Universal Robots PolyScope program: Renee_AI.urp

Program Renee_AI (installation=default directory=/ursim/programs createdIn=5.26.0 lastSavedIn=5.26.1 robotSerialNumber=20195599999)
Calibrated DH parameters: a=[0, -0.425, -0.3922, 0, 0, 0]; d=[0.1625, 0, 0, 0.1333, 0.0997, 0.0996]; alpha=[1.570796, 0, 0, 1.570796, -1.570796, 0]; deltaTheta=[0, 0, 0, 0, 0, 0]
InitVariablesNode
Robot Program (runOnlyOnce=true)
  var_1 := get_actual_tcp_pose()
  MoveJ speed 60 deg/s, acceleration 80 deg/s^2 (useActiveTCP=true optimoveEnabled=false optiMoveSpeed=0.3 optiMoveAcceleration=0.09) feature=Base
    Waypoint Variable (Variable): variable=var_1
  MoveJ speed 60 deg/s, acceleration 80 deg/s^2 (useActiveTCP=true positionType=JointAngles optimoveEnabled=false optiMoveSpeed=0.3 optiMoveAcceleration=0.09) feature=Base
    Waypoint Waypoint_1: TCP in base x=202.351 y=489.879 z=593.238 mm, rx=-1.5225 ry=0.5256 rz=-0.412 rad; joints [-127.677, -86.227, 99.579, -191.944, -86.567, 3.764] deg
  Script file /ursim/programs/generated_task.script
    | def inspection_program():
    |   # T_base_cam as a UR pose (position + axis-angle rotation vector)
    |   # Derived from the 4x4 transformation matrix T_base_cam
    |   global T_base_cam = p[0.352728458264352, -0.21258760881184183, 0.11788934094986696, -1.538543, 0.024168, 0.017202]
    | 
    |   # Offset to apply in camera frame: -0.4 m in camera X
    |   global x_offset = -0.40
    | 
    |   # Movement parameters (conservative for inspection)
    |   global accel = 0.3
    |   global vel = 0.05
    | 
    |   # Compute the first waypoint pose
    |   local first_wp = pose_trans(T_base_cam, p[0.335 + x_offset, 0.143, 0.57, 0, 0, 0])
    | 
    |   # Use movej to safely approach the first waypoint (avoids protective stop)
    |   movej(first_wp, a=1.0, v=0.5)
    |   sleep(1.0)
    | 
    |   # --- Waypoint 2: top_tube_front ---
    |   movel(pose_trans(T_base_cam, p[0.381 + x_offset, 0.116, 0.57, 0, 0, 0]), a=accel, v=vel)
    |   sleep(1.0)
    | 
    |   # --- Waypoint 3: top_tube_rear ---
    |   movel(pose_trans(T_base_cam, p[0.65 + x_offset, 0.131, 0.57, 0, 0, 0]), a=accel, v=vel)
    |   sleep(1.0)
    | 
    |   # --- Waypoint 4: seat_post_clamp ---
    |   movel(pose_trans(T_base_cam, p[0.68 + x_offset, 0.11, 0.57, 0, 0, 0]), a=accel, v=vel)
    |   sleep(1.0)
    | 
    |   # --- Waypoint 5: seat_tube_lower ---
    |   movel(pose_trans(T_base_cam, p[0.627 + x_offset, 0.462, 0.57, 0, 0, 0]), a=accel, v=vel)
    |   sleep(1.0)
    | 
    |   # --- Waypoint 6: bottom_bracket ---
    |   movel(pose_trans(T_base_cam, p[0.615 + x_offset, 0.609, 0.57, 0, 0, 0]), a=accel, v=vel)
    |   sleep(1.0)
    | 
    |   # --- Waypoint 7: chainstay_front ---
    |   movel(pose_trans(T_base_cam, p[0.701 + x_offset, 0.609, 0.57, 0, 0, 0]), a=accel, v=vel)
    |   sleep(1.0)
    | 
    |   # --- Waypoint 8: rear_dropout ---
    |   movel(pose_trans(T_base_cam, p[0.888 + x_offset, 0.586, 0.57, 0, 0, 0]), a=accel, v=vel)
    |   sleep(1.0)
    | 
    |   # --- Waypoint 9: seatstay_upper ---
    |   movel(pose_trans(T_base_cam, p[0.736 + x_offset, 0.308, 0.57, 0, 0, 0]), a=accel, v=vel)
    |   sleep(1.0)
    | 
    |   # --- Waypoint 10: seat_post_clamp ---
    |   movel(pose_trans(T_base_cam, p[0.68 + x_offset, 0.131, 0.57, 0, 0, 0]), a=accel, v=vel)
    |   sleep(1.0)
    | 
    |   # --- Waypoint 11: top_tube_rear ---
    |   movel(pose_trans(T_base_cam, p[0.65 + x_offset, 0.131, 0.57, 0, 0, 0]), a=accel, v=vel)
    |   sleep(1.0)
    | 
    |   # --- Waypoint 12: top_tube_front ---
    |   movel(pose_trans(T_base_cam, p[0.381 + x_offset, 0.116, 0.57, 0, 0, 0]), a=accel, v=vel)
    |   sleep(1.0)
    | 
    |   # --- Waypoint 13: head_tube ---
    |   movel(pose_trans(T_base_cam, p[0.335 + x_offset, 0.143, 0.57, 0, 0, 0]), a=accel, v=vel)
    |   sleep(1.0)
    | 
    |   # --- Waypoint 14: down_tube_upper ---
    |   movel(pose_trans(T_base_cam, p[0.355 + x_offset, 0.256, 0.57, 0, 0, 0]), a=accel, v=vel)
    |   sleep(1.0)
    | 
    |   # --- Waypoint 15: down_tube_lower ---
    |   movel(pose_trans(T_base_cam, p[0.545 + x_offset, 0.591, 0.57, 0, 0, 0]), a=accel, v=vel)
    |   sleep(1.0)
    | 
    |   # --- Waypoint 16: bottom_bracket ---
    |   movel(pose_trans(T_base_cam, p[0.615 + x_offset, 0.609, 0.57, 0, 0, 0]), a=accel, v=vel)
    |   sleep(1.0)
    | 
    | end
    | inspection_program()
